Universal Robots URScript: T015_codellama_34b_baseline_rep1.urscript

def program():
    # Home the robot
    movej(p[0, 0, 0, 0, 0, 0], v=350.0)

    # Move above the marking surface
    movel(p[0, 0, 100, 0, 0, 0], v=300.0)

    # Descend
